TYPE ST_Pick :
STRUCT
	bActive		: BOOL;		// 고른 값이 있음
	fValue		: REAL;		// kW 또는 kvar
	nModule		: UINT;		// 고른 지령원 모듈 ID
	bNew		: BOOL;		// 고른 지령원이 이번 스캔에 새 지령을 냄
END_STRUCT
END_TYPE

(* stored: Version 1.1.0.1, ProductVersion 3.1.4024.15
   DUT ST_Pick: Id {8b27862f-835e-4a01-b272-507e93468bb2} *)
